(*
SPDX-FileCopyrightText: © 2026 Oleksandr Tiutyk <trofimich@gmail.com>
SPDX-License-Identifier: MIT
License: https://opensource.org/license/mit
*)

(*!
<summary>Provides fluent assertions on a copied LTIME_OF_DAY value.</summary>
<description>
Copies actual into persistent instance storage before the entry method returns; literals and expression
results therefore remain valid throughout the immediate chain. Owns no heap allocation or pointed-to resource.
The message prefixes every failure until the next preparation. Finish one chain before starting another on
the owning Assertions provider. Use only from the owning test callback on one task, without reentry.
Obtain this context from the owning provider; direct unprepared use is unsupported.
Expected arguments use the declared IEC type; ordinary compiler conversions happen before comparison.
This context does not depend on another assertion context.
Object metadata is available before preparation; inherited equality compares instance identity.
Ordering uses the native IEC comparison of time since midnight, without a duration conversion or wrap-around.
</description>
*)

{attribute 'no_explicit_call' := 'do not call this function block directly'}
FUNCTION_BLOCK LongTimeOfDayAssertionContext EXTENDS TOF_Core.Object
VAR_STAT
	{attribute 'hide'}
	_ClassName : STRING := __POUNAME();
END_VAR
VAR
	_Actual : LTIME_OF_DAY;
	_TestCase : ITestCase;
	_Message : WSTRING(255);
END_VAR

(*!
<summary>Provides the implementation class name.</summary>
<description>
Borrowed read-only reference to compiler-initialized storage, valid throughout the instance lifetime.
Do not modify the returned reference; no ownership is transferred.
</description>
*)
{attribute 'monitoring' := 'call'}
PROPERTY ClassName : REFERENCE TO STRING
GET
ClassName REF= _ClassName;
END_GET
END_PROPERTY

(*!
<summary>Asserts that the actual value is strictly greater than expected.</summary>
<description>
Records failure without interrupting the callback; preserves the message for the rest of the chain.
</description>
<param name="expected">Expected value converted by the compiler to LTIME_OF_DAY.</param>
*)
METHOD FINAL IsGreaterThan : REFERENCE TO LongTimeOfDayAssertionContext
VAR_INPUT
	expected : LTIME_OF_DAY;
END_VAR
IF _Actual <= expected THEN
	failComparison(
		expected := expected,
		expectation := "Expected value > "
	);
END_IF

IsGreaterThan REF= THIS^;
END_METHOD

(*!
<summary>Asserts that the actual value meets the inclusive lower boundary.</summary>
<description>
Records failure without interrupting the callback; preserves the message for the rest of the chain.
</description>
<param name="expected">Expected value converted by the compiler to LTIME_OF_DAY.</param>
*)
METHOD FINAL IsGreaterThanOrEquals : REFERENCE TO LongTimeOfDayAssertionContext
VAR_INPUT
	expected : LTIME_OF_DAY;
END_VAR
IF _Actual < expected THEN
	failComparison(
		expected := expected,
		expectation := "Expected value >= "
	);
END_IF

IsGreaterThanOrEquals REF= THIS^;
END_METHOD

(*!
<summary>Asserts that the actual value is strictly less than expected.</summary>
<description>
Records failure without interrupting the callback; preserves the message for the rest of the chain.
</description>
<param name="expected">Expected value converted by the compiler to LTIME_OF_DAY.</param>
*)
METHOD FINAL IsLessThan : REFERENCE TO LongTimeOfDayAssertionContext
VAR_INPUT
	expected : LTIME_OF_DAY;
END_VAR
IF _Actual >= expected THEN
	failComparison(
		expected := expected,
		expectation := "Expected value < "
	);
END_IF

IsLessThan REF= THIS^;
END_METHOD

(*!
<summary>Asserts that the actual value meets the inclusive upper boundary.</summary>
<description>
Records failure without interrupting the callback; preserves the message for the rest of the chain.
</description>
<param name="expected">Expected value converted by the compiler to LTIME_OF_DAY.</param>
*)
METHOD FINAL IsLessThanOrEquals : REFERENCE TO LongTimeOfDayAssertionContext
VAR_INPUT
	expected : LTIME_OF_DAY;
END_VAR
IF _Actual > expected THEN
	failComparison(
		expected := expected,
		expectation := "Expected value <= "
	);
END_IF

IsLessThanOrEquals REF= THIS^;
END_METHOD

(*!
<summary>Provides the library namespace.</summary>
<description>
Borrowed read-only reference to the compiler-initialized namespace, valid throughout the instance lifetime.
Do not modify the returned reference; no ownership is transferred.
</description>
*)
{attribute 'monitoring' := 'call'}
PROPERTY NamespaceName : REFERENCE TO STRING
GET
NamespaceName REF= CurrentNamespace.Name;
END_GET
END_PROPERTY

(*!
<summary>Asserts inequality with the expected value.</summary>
<description>
Records failure without interrupting the callback; preserves the message for the rest of the chain.
</description>
<param name="expected">Expected value converted by the compiler to LTIME_OF_DAY.</param>
*)
METHOD FINAL NotToBe : REFERENCE TO LongTimeOfDayAssertionContext
VAR_INPUT
	expected : LTIME_OF_DAY;
END_VAR
IF _Actual = expected THEN
	failComparison(
		expected := expected,
		expectation := "Expected value not to be: "
	);
END_IF

NotToBe REF= THIS^;
END_METHOD

(*!
<summary>Copies the actual operand and replaces the chain-wide message.</summary>
<description>
Called by the owning Assertions provider after it verifies the running test case.
No pointer to this method's input storage is retained. The receiver is borrowed until the next preparation;
the owning provider keeps it alive throughout the immediate chain.
</description>
<param name="actual">Value copied into this context.</param>
<param name="testCase">Borrowed failure receiver for the immediate chain.</param>
<param name="message">Copied diagnostic prefix, including empty to clear the previous prefix.</param>
*)
METHOD INTERNAL FINAL Prepare
VAR_INPUT
	actual : LTIME_OF_DAY;
	testCase : ITestCase;
	message : WSTRING(255);
END_VAR
_Actual := actual;
_TestCase := testCase;
_Message := message;
END_METHOD

(*!
<summary>Reports the byte size of this concrete instance.</summary>
<description>
Includes inline fields and nested instances, but excludes separately allocated payloads.
Obtaining the size does not transfer ownership or validate an arbitrary address.
</description>
*)
{attribute 'monitoring' := 'call'}
PROPERTY SelfSize : ULINT
GET
SelfSize := XSIZEOF(THIS^);
END_GET
END_PROPERTY

(*!
<summary>Asserts equality with the expected value.</summary>
<description>
Records failure without interrupting the callback; preserves the message for the rest of the chain.
</description>
<param name="expected">Expected value converted by the compiler to LTIME_OF_DAY.</param>
*)
METHOD FINAL ToBe : REFERENCE TO LongTimeOfDayAssertionContext
VAR_INPUT
	expected : LTIME_OF_DAY;
END_VAR
IF _Actual <> expected THEN
	failComparison(
		expected := expected,
		expectation := "Expected: "
	);
END_IF

ToBe REF= THIS^;
END_METHOD

(*!
<summary>Formats a failed typed predicate and reports it with the chain message.</summary>
<description>
Does not change operands or chain state. The receiver retains its first failure. Reporting exceptions
propagate to the enclosing test callback handler; an unprepared receiver is a configuration error.
</description>
<param name="expected">Typed expected operand used only for this diagnostic.</param>
<param name="expectation">Prefix identifying the failed predicate.</param>
*)
METHOD PRIVATE failComparison
VAR_INPUT
	expected : LTIME_OF_DAY;
	expectation : WSTRING(40);
END_VAR
VAR
	actualText : WSTRING(255);
	expectedText : WSTRING(255);
	diagnostic : TOF_Core.ERROR_MESSAGE;
END_VAR
actualText := TO_WSTRING(_Actual);
expectedText := TO_WSTRING(expected);

diagnostic := TOF_Core.WideStrings.Concat255(
	expectation,
	expectedText,
	", but was: ",
	actualText
);

TestServices.ReportAssertionFailure(
	testCase := _TestCase,
	message := _Message,
	sourceClassName := ClassName,
	defaultMessage := diagnostic
);
END_METHOD

END_FUNCTION_BLOCK

(* stored: Version 1.1.0.1
   POU LongTimeOfDayAssertionContext: Id {07b25ffc-0dd3-4d40-93eb-31722f786696}, SpecialFunc None
   Folder Service methods: Id {e0f705e2-2f35-4d1c-887d-2c65eba43693}
   Property ClassName: Id {dc1a19a1-f2fc-4211-abe4-c703a362dfd9}
   Get Get: Id {a771c455-285f-45e4-896b-8c998e19f9c0}
   Method IsGreaterThan: Id {e8549bcf-9443-4116-9850-79ffbf968301}
   Method IsGreaterThanOrEquals: Id {47606ffc-1b27-4431-9ba1-5b04a895b4a3}
   Method IsLessThan: Id {417ca762-a3aa-4005-bc5b-ace3edc06ff2}
   Method IsLessThanOrEquals: Id {186e1d72-33ae-4b7f-9bfd-d66e1a9ff843}
   Property NamespaceName: Id {3be9de72-135a-4302-80e9-0d202f4b29be}
   Get Get: Id {b38ffcb2-f716-458e-a795-c04bb48809cd}
   Method NotToBe: Id {77b25070-b9e6-4ab4-9c22-8928ea727881}
   Method Prepare: Id {3ad52fd9-ae8e-4710-9941-ec0f38ba4de0}
   Property SelfSize: Id {3765c2fe-cfd9-48c5-bd9e-525123f447ee}
   Get Get: Id {b851f4e9-0e49-4bc5-be5f-59ece0ee51a3}
   Method ToBe: Id {4e64f39c-51a3-419c-9a60-7ce5e04c7960}
   Method failComparison: Id {0adc249e-28a5-4217-b4fd-99cd7fb9faea} *)
